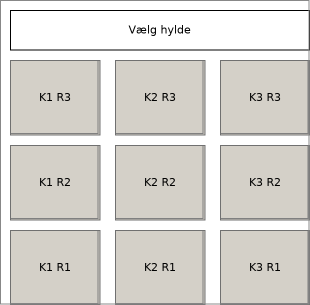
VISUALIZATION VisuShelf  // 310x305
    Rectangle (10,10 300x40), "Vælg hylde"
    Button (10,60 90x75), "K1 R3"
        OnMouseClick: execute {
            MAIN.nSelColumn := 1;
            MAIN.nSelRow := 3;
            MAIN.bShelfSelected := TRUE;
        }
    Button (115,60 90x75), "K2 R3"
        OnMouseClick: execute {
            MAIN.nSelColumn := 2;
            MAIN.nSelRow := 3;
            MAIN.bShelfSelected := TRUE;
        }
    Button (220,60 90x75), "K3 R3"
        OnMouseClick: execute {
            MAIN.nSelColumn := 3;
            MAIN.nSelRow := 3;
            MAIN.bShelfSelected := TRUE;
        }
    Button (10,145 90x75), "K1 R2"
        OnMouseClick: execute {
            MAIN.nSelColumn := 1;
            MAIN.nSelRow := 2;
            MAIN.bShelfSelected := TRUE;
        }
    Button (115,145 90x75), "K2 R2"
        OnMouseClick: execute {
            MAIN.nSelColumn := 2;
            MAIN.nSelRow := 2;
            MAIN.bShelfSelected := TRUE;
        }
    Button (220,145 90x75), "K3 R2"
        OnMouseClick: execute {
            MAIN.nSelColumn := 3;
            MAIN.nSelRow := 2;
            MAIN.bShelfSelected := TRUE;
        }
    Button (10,230 90x75), "K1 R1"
        OnMouseClick: execute {
            MAIN.nSelColumn := 1;
            MAIN.nSelRow := 1;
            MAIN.bShelfSelected := TRUE;
        }
    Button (115,230 90x75), "K2 R1"
        OnMouseClick: execute {
            MAIN.nSelColumn := 2;
            MAIN.nSelRow := 1;
            MAIN.bShelfSelected := TRUE;
        }
    Button (220,230 90x75), "K3 R1"
        OnMouseClick: execute {
            MAIN.nSelColumn := 3;
            MAIN.nSelRow := 1;
            MAIN.bShelfSelected := TRUE;
        }
END_VISUALIZATION

(* stored: Version 1.1.0.1, ProductVersion 3.1.4024.12
   Visu VisuShelf: Id {4d892f42-4e76-41ef-8cca-c48c99f8196c} *)
